Staubli VAL3: insertItem.pgx

public program insertItem(string x_sKey, string& x_sIndex, string x_sTRAJname, num x_nType, bool& x_bToSave)
  local num l_nIndex
  local bool l_bResult
  local num l_i
begin
  if x_sIndex!=""
    toNum(x_sIndex,l_nIndex,l_bResult)
    if l_bResult
      if l_nIndex==0 and progTemp:pProgItem[x_sKey].pProgTemplate[l_nIndex].sTRAJname==""
        progTemp:pProgItem[x_sKey].pProgTemplate[l_nIndex].sTRAJname=x_sTRAJname
        progTemp:pProgItem[x_sKey].pProgTemplate[l_nIndex].nType=x_nType
      else
        // l_nIndex=l_nIndex+1
        //insert(progTemp:pProgItem[x_sKey].pProgTemplate[l_nIndex])
        //l_nIndex=x_nIndex+1
        //insert(progTemp:pProgItem[x_sKey].pProgTemplate[x_nIndex+1])
        append(progTemp:pProgItem[x_sKey].pProgTemplate)
        for l_i = size(progTemp:pProgItem[x_sKey].pProgTemplate)-1 to l_nIndex step -1
          call copyPara(x_sKey,l_i-1,l_i)
        endFor
        progTemp:pProgItem[x_sKey].pProgTemplate[l_nIndex].sTRAJname=x_sTRAJname
        progTemp:pProgItem[x_sKey].pProgTemplate[l_nIndex].nType=x_nType
      endIf
      switch x_nType
        case 0
          x_sIndex=toString("",l_nIndex)+",TRAJ->"+x_sTRAJname
        break
        case 1
          x_sIndex=toString("",l_nIndex)+",ACTION->"+x_sTRAJname
        break
        case 2
          x_sIndex=toString("",l_nIndex)+",PROG->"+x_sTRAJname
        break
      endSwitch

      x_bToSave=true
    endIf
  else
    userPageAlert("未选中项目！")
  endIf
end
